// TIA Portal project "SmartFactory_FactoryIO_SortingStation" (V20)

(* hardware
DEVICE "S71500/ET200MP-Station_1"  S7-1500 station
   slot 0: "."  Rack  6ES7 590-1***0-0AA0
   slot 1: "PLC_1"  CPU 1511-1 PN  6ES7 511-1AK02-0AB0  V2.9
      slot 3: "CPU-Display_1"  6ES7591-1AA00-0AA0
      slot 32768: "PLC"  X1
         slot 32769: "Port_1"  X1 P1
         slot 32770: "Port_2"  X1 P2
      slot 34817: "Virtual CP interface port_1"  Virtual CP interface port  Virtual CP interface port
   slot 2: "AI 8xU/I/RTD/TC ST_1"  AI 8xU/I/RTD/TC ST  6ES7 531-7KF00-0AB0  V2.0
   slot 3: "AI 8xU/I/RTD/TC ST_2"  AI 8xU/I/RTD/TC ST  6ES7 531-7KF00-0AB0  V2.0
   slot 4: "AI 8xU/I/RTD/TC ST_3"  AI 8xU/I/RTD/TC ST  6ES7 531-7KF00-0AB0  V2.0
   slot 5: "AI 8xU/I/RTD/TC ST_4"  AI 8xU/I/RTD/TC ST  6ES7 531-7KF00-0AB0  V2.0
   slot 6: "DI 16x24VDC BA_1"  DI 16x24VDC BA  6ES7 521-1BH10-0AA0  V1.0
*)

// ===== PLC "PLC_1"  CPU 1511-1 PN =====

VAR_GLOBAL   // PLC tag table "Standard-Variablentabelle"
   "Start" AT %I0.0 : Bool;
   "Pause & Unpause" AT %I0.1 : Bool;
   "Reset" AT %I0.2 : Bool;
   "Pusher 1 front" AT %I0.3 : Bool;
   "Pusher 2 front" AT %I0.4 : Bool;
   "Pusher 1 back" AT %I0.5 : Bool;
   "Pusher 2 back" AT %I0.6 : Bool;
   "At pusher 1 exit" AT %I0.7 : Bool;
   "At pusher 2 exit" AT %I1.0 : Bool;
   "Sensor 1" AT %I1.1 : Bool;
   "Sensor 2" AT %I1.2 : Bool;
   "Vision sensor 1" AT %ID30 : DInt;
   "Vision sensor 2" AT %ID34 : DInt;
   "Start light" AT %Q0.0 : Bool;
   "P & UP light" AT %Q0.1 : Bool;
   "Reset light" AT %Q0.2 : Bool;
   "Conveyor 1" AT %Q0.3 : Bool;
   "Conveyor 2" AT %Q0.4 : Bool;
   "Entry conveyor 1" AT %Q0.5 : Bool;
   "Entry conveyor 2" AT %Q0.6 : Bool;
   "Pusher 1" AT %Q0.7 : Bool;
   "Pusher 2" AT %Q1.0 : Bool;
   "Blue count" AT %QD30 : DInt;
   "Green count" AT %QD34 : DInt;
   "SYS_RUN_MEM" AT %M0.0 : Bool;
   "SYS_UNPAUSED_MEM" AT %M0.1 : Bool;
   "CASE_C1GREEN_C2BLUE" AT %M0.2 : Bool;
   "GB_ENTRY_CONV1_MEM" AT %M0.3 : Bool;
   "GB_SENSOR1_PULSE_C1" AT %M0.4 : Bool;
   "GB_SENSOR1_NEG_C1" AT %M0.5 : Bool;
   "GB_CONVEYOR1_MEM" AT %M0.6 : Bool;
   "GB_ENTRY_CONV2_MEM" AT %M1.0 : Bool;
   "GB_ATPUSHER2EXIT_NEG_C2" AT %M1.1 : Bool;
   "GB_CONVEYOR2_MEM" AT %M1.2 : Bool;
   "GB_SENSOR1_NEG_P1" AT %M1.3 : Bool;
   "GB_PUSHER1_MEM" AT %M1.4 : Bool;
   "GB_CASE_EXIT" AT %M1.5 : Bool;
   "GB_SENSOR1_NEG_EC1" AT %M1.6 : Bool;
   "GB_ATPUSHER2EXIT_NEG_EC1" AT %M0.7 : Bool;
   "CASE_C1BLUE_C2GREEN" AT %M1.7 : Bool;
   "CASE_BOTH_BLUE" AT %M2.0 : Bool;
   "CASE_BOTH_GREEN" AT %M2.1 : Bool;
   "BG_ENTRY_C1C2_MEM" AT %M2.2 : Bool;
   "BG_CASE_EXIT" AT %M2.3 : Bool;
   "CASE_GB_RESETS_BG_PULSE" AT %M2.4 : Bool;
   "CASE_BG_RESETS_GB_PULSE" AT %M2.5 : Bool;
   "CASE_BB_RESETS_GB_PULSE" AT %M2.6 : Bool;
   "CASE_GG_RESETS_GB_PULSE" AT %M2.7 : Bool;
   "CASE_BB_RESETS_BG_PULSE" AT %M3.0 : Bool;
   "CASE_GG_RESETS_BG_PULSE" AT %M3.1 : Bool;
   "CASE_GB_RESETS_BB_PULSE" AT %M3.2 : Bool;
   "CASE_BG_RESETS_BB_PULSE" AT %M3.3 : Bool;
   "CASE_GG_RESETS_BB_PULSE" AT %M3.4 : Bool;
   "BB_CASE_EXIT" AT %M3.5 : Bool;
   "BB_ENTRY_CONV1_MEM" AT %M3.6 : Bool;
   "BB_CONVEYOR1_MEM" AT %M3.7 : Bool;
   "BB_ENTRY_CONV2_MEM" AT %M4.0 : Bool;
   "BB_CONVEYOR2_MEM" AT %M4.1 : Bool;
   "BB_PUSHER2_MEM" AT %M4.2 : Bool;
   "BB_SENSOR2_NEG" AT %M4.3 : Bool;
   "BB_SENSOR2_PULSE" AT %M4.4 : Bool;
   "BB_SENSOR2_NEG_C2" AT %M4.5 : Bool;
   "BB_SENSOR2_NEG_P2" AT %M4.6 : Bool;
   "BB_ATPUSHER1EXIT_NEG" AT %M4.7 : Bool;
   "BB_ATPUSHER1EXIT_NEG_EC1" AT %M5.0 : Bool;
   "CASE_GB_RESETS_GG_PULSE" AT %M5.1 : Bool;
   "CASE_BG_RESETS_GG_PULSE" AT %M5.2 : Bool;
   "CASE_BB_RESETS_GG_PULSE" AT %M5.3 : Bool;
   "GG_ENTRY_CONV1_MEM" AT %M5.4 : Bool;
   "GG_CONVEYOR1_MEM" AT %M5.5 : Bool;
   "GG_ENTRY_CONV2_MEM" AT %M5.6 : Bool;
   "GG_CONVEYOR2_MEM" AT %M5.7 : Bool;
   "GG_PUSHER1_MEM" AT %M6.0 : Bool;
   "GG_SENSOR1_PULSE" AT %M6.1 : Bool;
   "GG_SENSOR1_NEG_EC1" AT %M6.2 : Bool;
   "GG_SENSOR1_NEG_C1" AT %M6.3 : Bool;
   "GG_SENSOR1_NEG_P1" AT %M6.4 : Bool;
   "GG_ATPUSHER2EXIT_NEG" AT %M6.5 : Bool;
   "GG_ATPUSHER2EXIT_NEG_EC1" AT %M6.6 : Bool;
   "BG_SENSOR1_PULSE" AT %M6.7 : Bool;
   "BG_CONV1CONV2_MEM" AT %M7.0 : Bool;
   "BG_SENSOR1_NEG" AT %M7.1 : Bool;
   "BG_ATPUSHER1EXIT_NEG_C1C2" AT %M7.2 : Bool;
   "BG_ATPUSHER1EXIT_NEG_EC1EC2" AT %M7.3 : Bool;
   "CNT_BLUE_TRIGGER" AT %M7.4 : Bool;
   "CNT_GREEN_TRIGGER" AT %M7.5 : Bool;
   "SYS_PAUSED_MEM" AT %M7.6 : Bool;
END_VAR

// folder: System blocks/Program resources

DATA_BLOCK "IEC_Counter_0_DB"   // DB1
{ S7_Optimized_Access := 'TRUE' }
AUTHOR : SIMATIC
FAMILY : IEC
NAME : DCNTR
VERSION : 1.2
// stored: InstanceOfName IEC_DCOUNTER
"IEC_DCOUNTER"
BEGIN
END_DATA_BLOCK

DATA_BLOCK "IEC_Counter_0_DB_1"   // DB2
{ S7_Optimized_Access := 'TRUE' }
AUTHOR : SIMATIC
FAMILY : IEC
NAME : DCNTR
VERSION : 1.2
// stored: InstanceOfName IEC_DCOUNTER
"IEC_DCOUNTER"
BEGIN
END_DATA_BLOCK

// folder: (top level)

FUNCTION "MHJ-PLC-Lab-Function-S71500" : Void   // FC9000, SCL
{ S7_Optimized_Access := 'TRUE' }
VERSION : 0.1
   VAR_TEMP
      Value : Byte;
      ForCounter : Int;
   END_VAR
   VAR CONSTANT
      Value_01_DW : DWord := 16#1223_5486;
      Value_02_DW : DWord := 16#A6C9_D1F5;
   END_VAR
BEGIN

   #Value:=PEEK(area := 16#82,
        dbNumber := 0,
        byteOffset := 511);
   #Value := #Value + 1;

   POKE(area := 16#82,
        dbNumber := 0,
        byteOffset := 511,
        value := #Value);

   POKE(area := 16#82,
        dbNumber := 0,
        byteOffset := 1016,
        value := #Value_01_DW);
   POKE(area := 16#82,
        dbNumber := 0,
        byteOffset := 1020,
        value := #Value_02_DW);

   FOR #ForCounter := 0 TO 63 DO
       #Value:=PEEK(area := 16#1,
            dbNumber := 0,
            byteOffset := #ForCounter);
       POKE(area := 16#81,
            dbNumber := 0,
            byteOffset := #ForCounter,
            value := #Value);
   END_FOR;
   #Value := PEEK(area := 16#1,
                  dbNumber := 0,
                  byteOffset := 512);
   POKE(area := 16#82,
        dbNumber := 0,
        byteOffset := 512,
        value := #Value);
END_FUNCTION

ORGANIZATION_BLOCK "Main"   // OB1, LAD, ProgramCycle
TITLE = "Main Program Sweep (Cycle)"
{ S7_Optimized_Access := 'TRUE' }
VERSION : 0.1
   VAR_INPUT
      Initial_Call : Bool;   // Initial call of this OB
      Remanence : Bool;   // =True, if remanent data are available
   END_VAR
   VAR_TEMP   // added for the SCL form of the ladder/FBD networks
      _w1 : Bool;
      _w2 : Bool;
      _w3 : Bool;
      _w4 : Bool;
      _w5 : Bool;
      _w6 : Bool;
      _w7 : Bool;
      _w8 : Bool;
      _w9 : Bool;
      _w10 : Bool;
      _w11 : Bool;
      _w12 : Bool;
      _w13 : Bool;
      _w14 : Bool;
   END_VAR
BEGIN

REGION Network 1
   // Lien TIA ↔ Factory I/O (FC9000), ne pas supprimer.
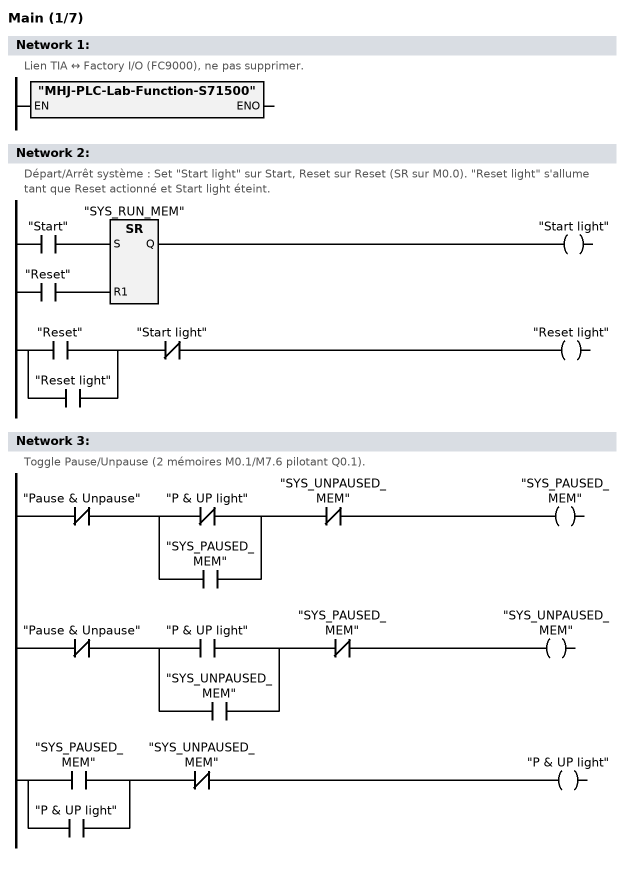
   RUNG wire#powerrail
      "MHJ-PLC-Lab-Function-S71500"()
   END_RUNG
   // the same network as SCL:
   "MHJ-PLC-Lab-Function-S71500"();
END_REGION

REGION Network 2
   // Départ/Arrêt système : Set "Start light" sur Start, Reset sur Reset (SR sur M0.0). "Reset light" s'allume tant que Reset actionné et Start light éteint.
   RUNG wire#powerrail
      Contact( "Start" )
      S_SR(operand := "SYS_RUN_MEM", r1 := wire#w1)
      Coil( "Start light" )
   END_RUNG
   RUNG wire#powerrail
      Contact( "Reset" )
   END_RUNG wire#w1
   RUNG wire#powerrail
      Contact( "Reset" )
      wire#w2
      I_Contact( "Start light" )
      Coil( "Reset light" )
   END_RUNG
   RUNG wire#powerrail
      Contact( "Reset light" )
   END_RUNG wire#w2
   // the same network as SCL:
   IF "Start" THEN
       "SYS_RUN_MEM" := TRUE;   // SR flip-flop
   END_IF;
   IF "Reset" THEN "SYS_RUN_MEM" := FALSE; END_IF;
   "Start light" := "SYS_RUN_MEM";
   "Reset light" := ("Reset" OR "Reset light") AND NOT "Start light";
END_REGION

REGION Network 3
   // Toggle Pause/Unpause (2 mémoires M0.1/M7.6 pilotant Q0.1).
   RUNG wire#powerrail
      I_Contact( "Pause & Unpause" )
      wire#w1
      I_Contact( "P & UP light" )
      wire#w2
      I_Contact( "SYS_UNPAUSED_MEM" )
      Coil( "SYS_PAUSED_MEM" )
   END_RUNG
   RUNG wire#w1
      Contact( "SYS_PAUSED_MEM" )
   END_RUNG wire#w2
   RUNG wire#powerrail
      I_Contact( "Pause & Unpause" )
      wire#w3
      Contact( "P & UP light" )
      wire#w4
      I_Contact( "SYS_PAUSED_MEM" )
      Coil( "SYS_UNPAUSED_MEM" )
   END_RUNG
   RUNG wire#w3
      Contact( "SYS_UNPAUSED_MEM" )
   END_RUNG wire#w4
   RUNG wire#powerrail
      Contact( "SYS_PAUSED_MEM" )
      wire#w5
      I_Contact( "SYS_UNPAUSED_MEM" )
      Coil( "P & UP light" )
   END_RUNG
   RUNG wire#powerrail
      Contact( "P & UP light" )
   END_RUNG wire#w5
   // the same network as SCL:
   "SYS_PAUSED_MEM" := NOT "Pause & Unpause" AND (NOT "P & UP light" OR "SYS_PAUSED_MEM") AND NOT "SYS_UNPAUSED_MEM";
   "SYS_UNPAUSED_MEM" := NOT "Pause & Unpause" AND ("P & UP light" OR "SYS_UNPAUSED_MEM") AND NOT "SYS_PAUSED_MEM";
   "P & UP light" := ("SYS_PAUSED_MEM" OR "P & UP light") AND NOT "SYS_UNPAUSED_MEM";
END_REGION

REGION Network 4
   // Détection de la combinaison couleur des 2 postes (Vision sensor 1=Bleu(1)/Vert(4), idem sensor 2). 4 cas mutuellement exclusifs mémorisés en SR, avec reset croisé par front montant dès qu'un autre cas se déclenche. Comptage Bleu/Vert en sortie (CTU sur "At pusher 1/2 exit").
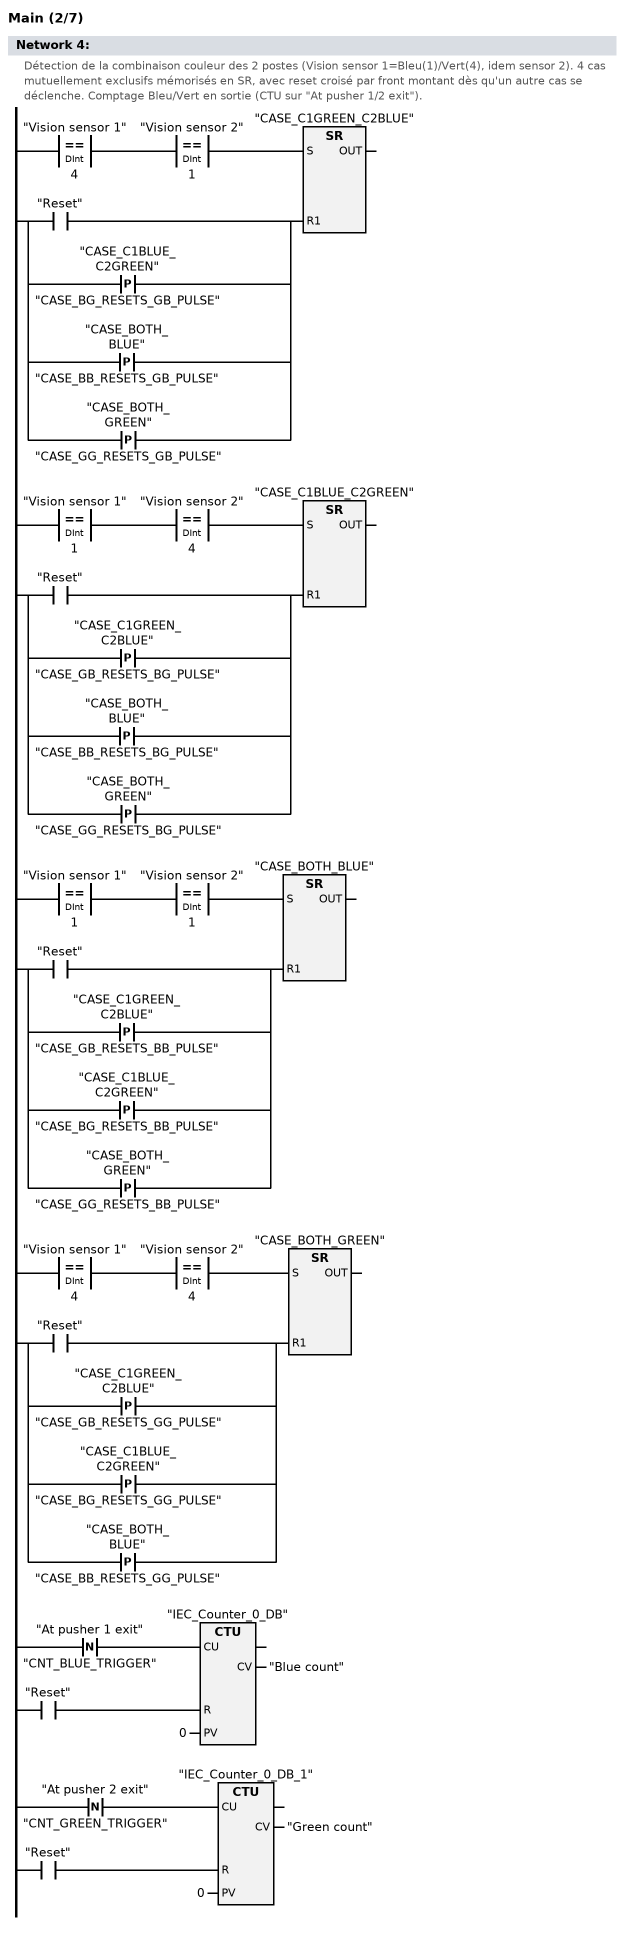
   #_w1 := "CASE_C1BLUE_C2GREEN" AND NOT "CASE_BG_RESETS_GB_PULSE";   // rising edge of "CASE_C1BLUE_C2GREEN"
   "CASE_BG_RESETS_GB_PULSE" := "CASE_C1BLUE_C2GREEN";
   #_w2 := "CASE_BOTH_BLUE" AND NOT "CASE_BB_RESETS_GB_PULSE";   // rising edge of "CASE_BOTH_BLUE"
   "CASE_BB_RESETS_GB_PULSE" := "CASE_BOTH_BLUE";
   #_w3 := "CASE_BOTH_GREEN" AND NOT "CASE_GG_RESETS_GB_PULSE";   // rising edge of "CASE_BOTH_GREEN"
   "CASE_GG_RESETS_GB_PULSE" := "CASE_BOTH_GREEN";
   IF ("Vision sensor 1" = 4) AND ("Vision sensor 2" = 1) THEN
       "CASE_C1GREEN_C2BLUE" := TRUE;   // SR flip-flop
   END_IF;
   IF "Reset" OR #_w1 OR #_w2 OR #_w3 THEN "CASE_C1GREEN_C2BLUE" := FALSE; END_IF;
   #_w4 := "CASE_C1GREEN_C2BLUE" AND NOT "CASE_GB_RESETS_BG_PULSE";   // rising edge of "CASE_C1GREEN_C2BLUE"
   "CASE_GB_RESETS_BG_PULSE" := "CASE_C1GREEN_C2BLUE";
   #_w5 := "CASE_BOTH_BLUE" AND NOT "CASE_BB_RESETS_BG_PULSE";   // rising edge of "CASE_BOTH_BLUE"
   "CASE_BB_RESETS_BG_PULSE" := "CASE_BOTH_BLUE";
   #_w6 := "CASE_BOTH_GREEN" AND NOT "CASE_GG_RESETS_BG_PULSE";   // rising edge of "CASE_BOTH_GREEN"
   "CASE_GG_RESETS_BG_PULSE" := "CASE_BOTH_GREEN";
   IF ("Vision sensor 1" = 1) AND ("Vision sensor 2" = 4) THEN
       "CASE_C1BLUE_C2GREEN" := TRUE;   // SR flip-flop
   END_IF;
   IF "Reset" OR #_w4 OR #_w5 OR #_w6 THEN "CASE_C1BLUE_C2GREEN" := FALSE; END_IF;
   #_w7 := "CASE_C1GREEN_C2BLUE" AND NOT "CASE_GB_RESETS_BB_PULSE";   // rising edge of "CASE_C1GREEN_C2BLUE"
   "CASE_GB_RESETS_BB_PULSE" := "CASE_C1GREEN_C2BLUE";
   #_w8 := "CASE_C1BLUE_C2GREEN" AND NOT "CASE_BG_RESETS_BB_PULSE";   // rising edge of "CASE_C1BLUE_C2GREEN"
   "CASE_BG_RESETS_BB_PULSE" := "CASE_C1BLUE_C2GREEN";
   #_w9 := "CASE_BOTH_GREEN" AND NOT "CASE_GG_RESETS_BB_PULSE";   // rising edge of "CASE_BOTH_GREEN"
   "CASE_GG_RESETS_BB_PULSE" := "CASE_BOTH_GREEN";
   IF ("Vision sensor 1" = 1) AND ("Vision sensor 2" = 1) THEN
       "CASE_BOTH_BLUE" := TRUE;   // SR flip-flop
   END_IF;
   IF "Reset" OR #_w7 OR #_w8 OR #_w9 THEN "CASE_BOTH_BLUE" := FALSE; END_IF;
   #_w10 := "CASE_C1GREEN_C2BLUE" AND NOT "CASE_GB_RESETS_GG_PULSE";   // rising edge of "CASE_C1GREEN_C2BLUE"
   "CASE_GB_RESETS_GG_PULSE" := "CASE_C1GREEN_C2BLUE";
   #_w11 := "CASE_C1BLUE_C2GREEN" AND NOT "CASE_BG_RESETS_GG_PULSE";   // rising edge of "CASE_C1BLUE_C2GREEN"
   "CASE_BG_RESETS_GG_PULSE" := "CASE_C1BLUE_C2GREEN";
   #_w12 := "CASE_BOTH_BLUE" AND NOT "CASE_BB_RESETS_GG_PULSE";   // rising edge of "CASE_BOTH_BLUE"
   "CASE_BB_RESETS_GG_PULSE" := "CASE_BOTH_BLUE";
   IF ("Vision sensor 1" = 4) AND ("Vision sensor 2" = 4) THEN
       "CASE_BOTH_GREEN" := TRUE;   // SR flip-flop
   END_IF;
   IF "Reset" OR #_w10 OR #_w11 OR #_w12 THEN "CASE_BOTH_GREEN" := FALSE; END_IF;
   #_w13 := NOT "At pusher 1 exit" AND "CNT_BLUE_TRIGGER";   // falling edge of "At pusher 1 exit"
   "CNT_BLUE_TRIGGER" := "At pusher 1 exit";
   "IEC_Counter_0_DB".CTU(CU := #_w13, R := "Reset", PV := 0, CV => "Blue count");
   #_w14 := NOT "At pusher 2 exit" AND "CNT_GREEN_TRIGGER";   // falling edge of "At pusher 2 exit"
   "CNT_GREEN_TRIGGER" := "At pusher 2 exit";
   "IEC_Counter_0_DB_1".CTU(CU := #_w14, R := "Reset", PV := 0, CV => "Green count");
END_REGION

REGION Network 5
   // Si le cas "Vert sur Conv1 / Bleu sur Conv2" est actif → saut vers Network 9, les Networks 10 à 12 sont ignorés ce cycle.
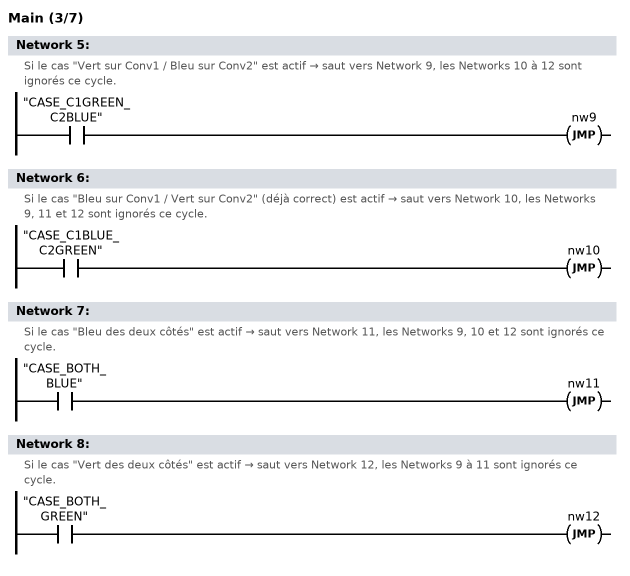
   RUNG wire#powerrail
      Contact( "CASE_C1GREEN_C2BLUE" )
      JumpCoil( nw9 )
   END_RUNG
   // the same network as SCL:
   IF "CASE_C1GREEN_C2BLUE" THEN GOTO nw9; END_IF;
END_REGION

REGION Network 6
   // Si le cas "Bleu sur Conv1 / Vert sur Conv2" (déjà correct) est actif → saut vers Network 10, les Networks 9, 11 et 12 sont ignorés ce cycle.
   RUNG wire#powerrail
      Contact( "CASE_C1BLUE_C2GREEN" )
      JumpCoil( nw10 )
   END_RUNG
   // the same network as SCL:
   IF "CASE_C1BLUE_C2GREEN" THEN GOTO nw10; END_IF;
END_REGION

REGION Network 7
   // Si le cas "Bleu des deux côtés" est actif → saut vers Network 11, les Networks 9, 10 et 12 sont ignorés ce cycle.
   RUNG wire#powerrail
      Contact( "CASE_BOTH_BLUE" )
      JumpCoil( nw11 )
   END_RUNG
   // the same network as SCL:
   IF "CASE_BOTH_BLUE" THEN GOTO nw11; END_IF;
END_REGION

REGION Network 8
   // Si le cas "Vert des deux côtés" est actif → saut vers Network 12, les Networks 9 à 11 sont ignorés ce cycle.
   RUNG wire#powerrail
      Contact( "CASE_BOTH_GREEN" )
      JumpCoil( nw12 )
   END_RUNG
   // the same network as SCL:
   IF "CASE_BOTH_GREEN" THEN GOTO nw12; END_IF;
END_REGION

REGION Network 9
   // Cas Vert/Bleu (positions inversées) : active les 2 convoyeurs d'entrée + convoyeur 1 sur détection Sensor 1, puis Pousseur 1 transfère l'objet Vert du convoyeur 1 vers le convoyeur 2 dès qu'il atteint la butée. RET dès que le cas GB n'est plus actif.
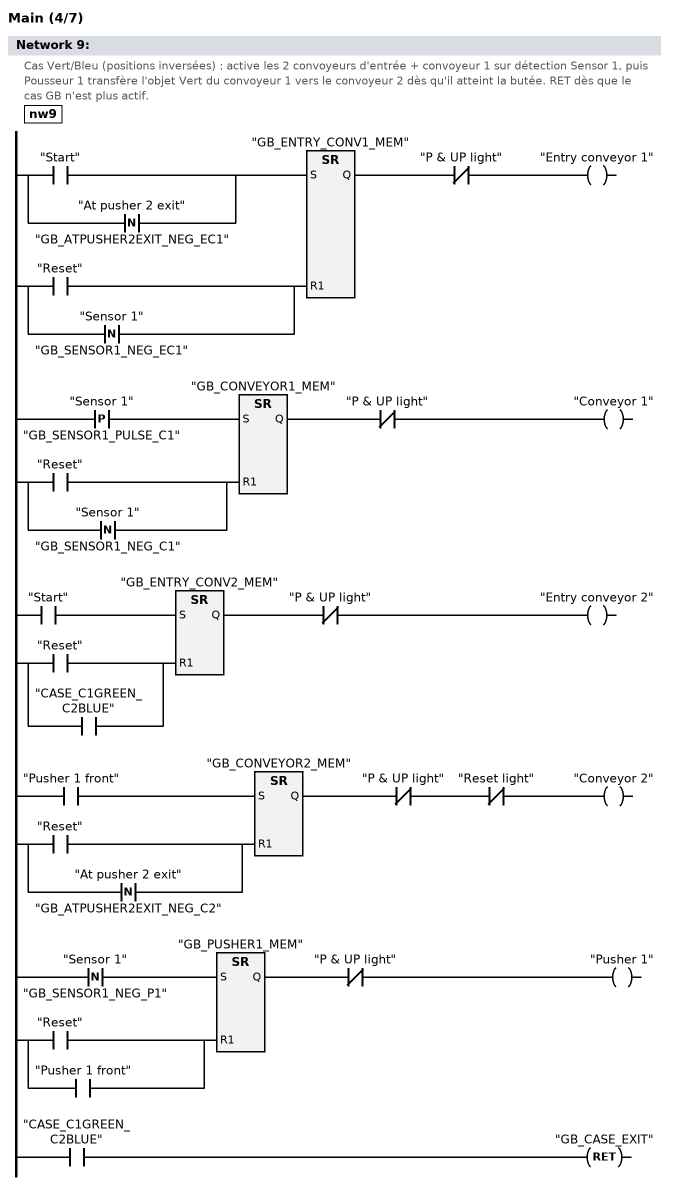
   nw9:
   #_w1 := NOT "At pusher 2 exit" AND "GB_ATPUSHER2EXIT_NEG_EC1";   // falling edge of "At pusher 2 exit"
   "GB_ATPUSHER2EXIT_NEG_EC1" := "At pusher 2 exit";
   #_w2 := NOT "Sensor 1" AND "GB_SENSOR1_NEG_EC1";   // falling edge of "Sensor 1"
   "GB_SENSOR1_NEG_EC1" := "Sensor 1";
   IF "Start" OR #_w1 THEN
       "GB_ENTRY_CONV1_MEM" := TRUE;   // SR flip-flop
   END_IF;
   IF "Reset" OR #_w2 THEN "GB_ENTRY_CONV1_MEM" := FALSE; END_IF;
   "Entry conveyor 1" := "GB_ENTRY_CONV1_MEM" AND NOT "P & UP light";
   #_w3 := "Sensor 1" AND NOT "GB_SENSOR1_PULSE_C1";   // rising edge of "Sensor 1"
   "GB_SENSOR1_PULSE_C1" := "Sensor 1";
   #_w4 := NOT "Sensor 1" AND "GB_SENSOR1_NEG_C1";   // falling edge of "Sensor 1"
   "GB_SENSOR1_NEG_C1" := "Sensor 1";
   IF #_w3 THEN
       "GB_CONVEYOR1_MEM" := TRUE;   // SR flip-flop
   END_IF;
   IF "Reset" OR #_w4 THEN "GB_CONVEYOR1_MEM" := FALSE; END_IF;
   "Conveyor 1" := "GB_CONVEYOR1_MEM" AND NOT "P & UP light";
   IF "Start" THEN
       "GB_ENTRY_CONV2_MEM" := TRUE;   // SR flip-flop
   END_IF;
   IF "Reset" OR "CASE_C1GREEN_C2BLUE" THEN "GB_ENTRY_CONV2_MEM" := FALSE; END_IF;
   "Entry conveyor 2" := "GB_ENTRY_CONV2_MEM" AND NOT "P & UP light";
   #_w5 := NOT "At pusher 2 exit" AND "GB_ATPUSHER2EXIT_NEG_C2";   // falling edge of "At pusher 2 exit"
   "GB_ATPUSHER2EXIT_NEG_C2" := "At pusher 2 exit";
   IF "Pusher 1 front" THEN
       "GB_CONVEYOR2_MEM" := TRUE;   // SR flip-flop
   END_IF;
   IF "Reset" OR #_w5 THEN "GB_CONVEYOR2_MEM" := FALSE; END_IF;
   "Conveyor 2" := "GB_CONVEYOR2_MEM" AND NOT "P & UP light" AND NOT "Reset light";
   #_w6 := NOT "Sensor 1" AND "GB_SENSOR1_NEG_P1";   // falling edge of "Sensor 1"
   "GB_SENSOR1_NEG_P1" := "Sensor 1";
   IF #_w6 THEN
       "GB_PUSHER1_MEM" := TRUE;   // SR flip-flop
   END_IF;
   IF "Reset" OR "Pusher 1 front" THEN "GB_PUSHER1_MEM" := FALSE; END_IF;
   "Pusher 1" := "GB_PUSHER1_MEM" AND NOT "P & UP light";
   IF "CASE_C1GREEN_C2BLUE" THEN
       ENO := "GB_CASE_EXIT";
       RETURN;
   END_IF;
END_REGION

REGION Network 10
   // Cas Bleu/Vert déjà en bonne position : active simplement les 2 convoyeurs d'entrée + les 2 convoyeurs principaux, aucun pousseur nécessaire.
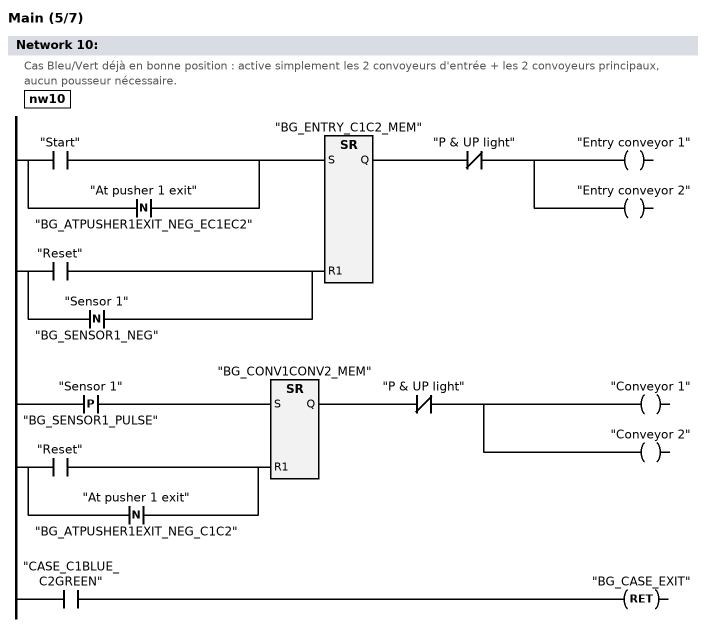
   nw10:
   #_w1 := NOT "At pusher 1 exit" AND "BG_ATPUSHER1EXIT_NEG_EC1EC2";   // falling edge of "At pusher 1 exit"
   "BG_ATPUSHER1EXIT_NEG_EC1EC2" := "At pusher 1 exit";
   #_w2 := NOT "Sensor 1" AND "BG_SENSOR1_NEG";   // falling edge of "Sensor 1"
   "BG_SENSOR1_NEG" := "Sensor 1";
   IF "Start" OR #_w1 THEN
       "BG_ENTRY_C1C2_MEM" := TRUE;   // SR flip-flop
   END_IF;
   IF "Reset" OR #_w2 THEN "BG_ENTRY_C1C2_MEM" := FALSE; END_IF;
   "Entry conveyor 1" := "BG_ENTRY_C1C2_MEM" AND NOT "P & UP light";
   "Entry conveyor 2" := "Entry conveyor 1";
   #_w3 := "Sensor 1" AND NOT "BG_SENSOR1_PULSE";   // rising edge of "Sensor 1"
   "BG_SENSOR1_PULSE" := "Sensor 1";
   #_w4 := NOT "At pusher 1 exit" AND "BG_ATPUSHER1EXIT_NEG_C1C2";   // falling edge of "At pusher 1 exit"
   "BG_ATPUSHER1EXIT_NEG_C1C2" := "At pusher 1 exit";
   IF #_w3 THEN
       "BG_CONV1CONV2_MEM" := TRUE;   // SR flip-flop
   END_IF;
   IF "Reset" OR #_w4 THEN "BG_CONV1CONV2_MEM" := FALSE; END_IF;
   "Conveyor 1" := "BG_CONV1CONV2_MEM" AND NOT "P & UP light";
   "Conveyor 2" := "Conveyor 1";
   IF "CASE_C1BLUE_C2GREEN" THEN
       ENO := "BG_CASE_EXIT";
       RETURN;
   END_IF;
END_REGION

REGION Network 11
   // Cas Bleu des deux côtés : Pousseur 2 renvoie l'objet Bleu en excès du convoyeur 2 vers le convoyeur 1 (symétrique de N9, sur Sensor 2/Pousseur 2).
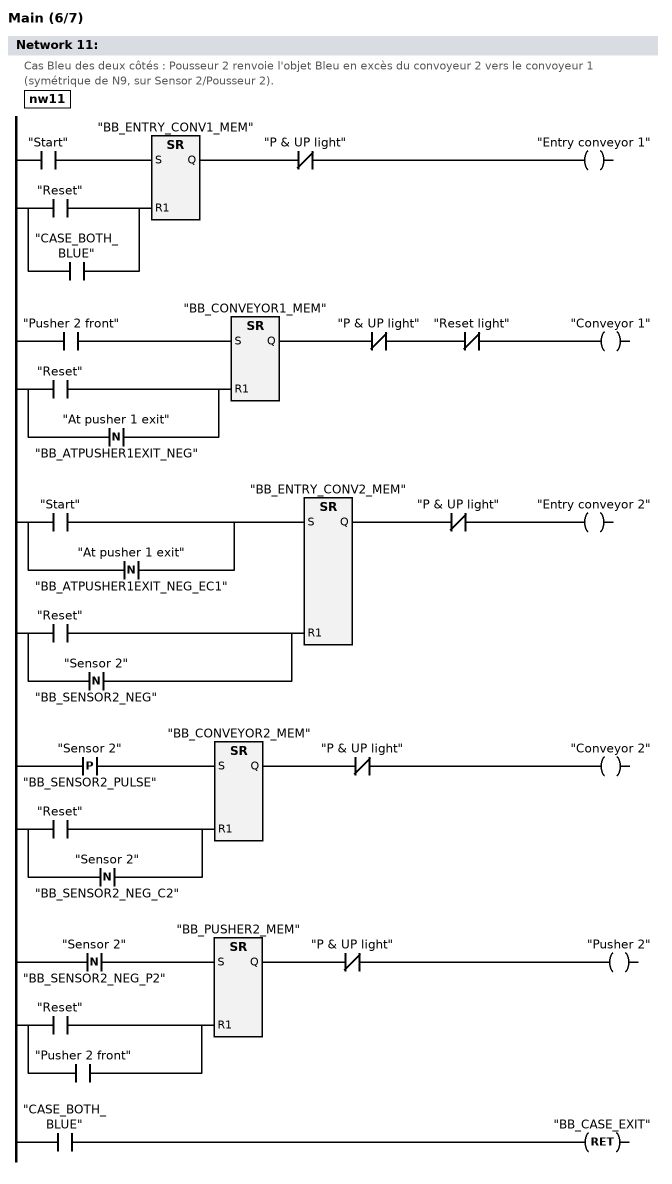
   nw11:
   IF "Start" THEN
       "BB_ENTRY_CONV1_MEM" := TRUE;   // SR flip-flop
   END_IF;
   IF "Reset" OR "CASE_BOTH_BLUE" THEN "BB_ENTRY_CONV1_MEM" := FALSE; END_IF;
   "Entry conveyor 1" := "BB_ENTRY_CONV1_MEM" AND NOT "P & UP light";
   #_w1 := NOT "At pusher 1 exit" AND "BB_ATPUSHER1EXIT_NEG";   // falling edge of "At pusher 1 exit"
   "BB_ATPUSHER1EXIT_NEG" := "At pusher 1 exit";
   IF "Pusher 2 front" THEN
       "BB_CONVEYOR1_MEM" := TRUE;   // SR flip-flop
   END_IF;
   IF "Reset" OR #_w1 THEN "BB_CONVEYOR1_MEM" := FALSE; END_IF;
   "Conveyor 1" := "BB_CONVEYOR1_MEM" AND NOT "P & UP light" AND NOT "Reset light";
   #_w2 := NOT "At pusher 1 exit" AND "BB_ATPUSHER1EXIT_NEG_EC1";   // falling edge of "At pusher 1 exit"
   "BB_ATPUSHER1EXIT_NEG_EC1" := "At pusher 1 exit";
   #_w3 := NOT "Sensor 2" AND "BB_SENSOR2_NEG";   // falling edge of "Sensor 2"
   "BB_SENSOR2_NEG" := "Sensor 2";
   IF "Start" OR #_w2 THEN
       "BB_ENTRY_CONV2_MEM" := TRUE;   // SR flip-flop
   END_IF;
   IF "Reset" OR #_w3 THEN "BB_ENTRY_CONV2_MEM" := FALSE; END_IF;
   "Entry conveyor 2" := "BB_ENTRY_CONV2_MEM" AND NOT "P & UP light";
   #_w4 := "Sensor 2" AND NOT "BB_SENSOR2_PULSE";   // rising edge of "Sensor 2"
   "BB_SENSOR2_PULSE" := "Sensor 2";
   #_w5 := NOT "Sensor 2" AND "BB_SENSOR2_NEG_C2";   // falling edge of "Sensor 2"
   "BB_SENSOR2_NEG_C2" := "Sensor 2";
   IF #_w4 THEN
       "BB_CONVEYOR2_MEM" := TRUE;   // SR flip-flop
   END_IF;
   IF "Reset" OR #_w5 THEN "BB_CONVEYOR2_MEM" := FALSE; END_IF;
   "Conveyor 2" := "BB_CONVEYOR2_MEM" AND NOT "P & UP light";
   #_w6 := NOT "Sensor 2" AND "BB_SENSOR2_NEG_P2";   // falling edge of "Sensor 2"
   "BB_SENSOR2_NEG_P2" := "Sensor 2";
   IF #_w6 THEN
       "BB_PUSHER2_MEM" := TRUE;   // SR flip-flop
   END_IF;
   IF "Reset" OR "Pusher 2 front" THEN "BB_PUSHER2_MEM" := FALSE; END_IF;
   "Pusher 2" := "BB_PUSHER2_MEM" AND NOT "P & UP light";
   IF "CASE_BOTH_BLUE" THEN
       ENO := "BB_CASE_EXIT";
       RETURN;
   END_IF;
END_REGION

REGION Network 12
   // Cas Vert des deux côtés : Pousseur 1 déplace l'objet Vert en excès du convoyeur 1 vers le convoyeur 2 (même logique que N9).
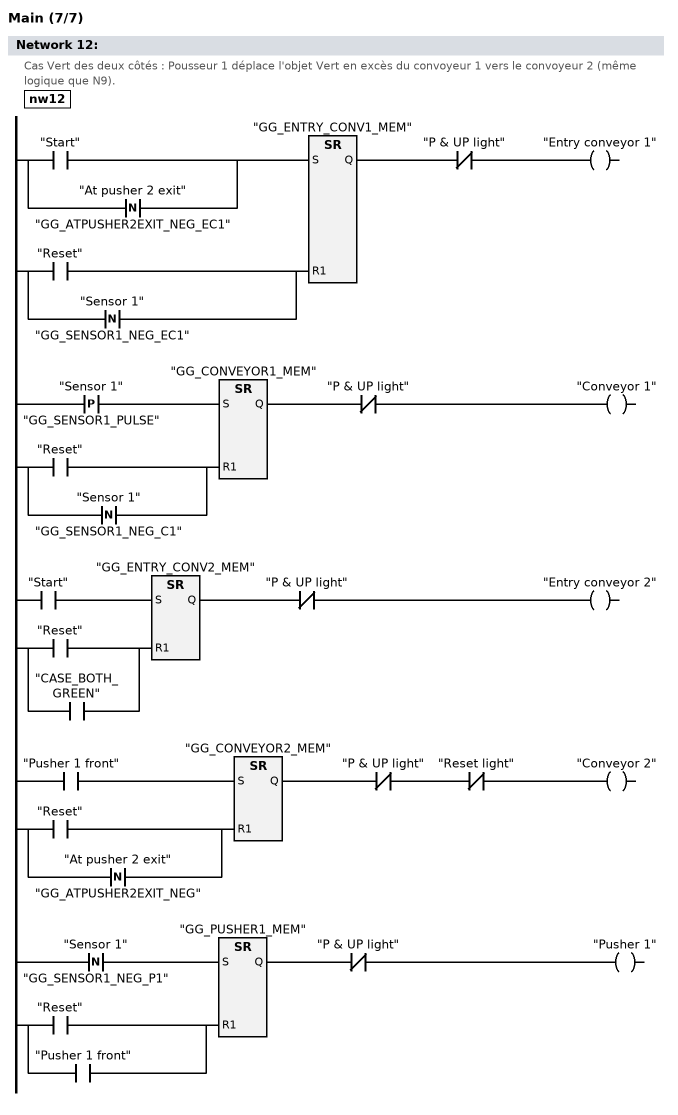
   Label( nw12 )
   RUNG wire#powerrail
      Contact( "Start" )
      wire#w1
      S_SR(operand := "GG_ENTRY_CONV1_MEM", r1 := wire#w2)
      I_Contact( "P & UP light" )
      Coil( "Entry conveyor 1" )
   END_RUNG
   RUNG wire#powerrail
      N_Contact(operand := "At pusher 2 exit", bit := "GG_ATPUSHER2EXIT_NEG_EC1")
   END_RUNG wire#w1
   RUNG wire#powerrail
      Contact( "Reset" )
   END_RUNG wire#w2
   RUNG wire#powerrail
      N_Contact(operand := "Sensor 1", bit := "GG_SENSOR1_NEG_EC1")
   END_RUNG wire#w2
   RUNG wire#powerrail
      P_Contact(operand := "Sensor 1", bit := "GG_SENSOR1_PULSE")
      S_SR(operand := "GG_CONVEYOR1_MEM", r1 := wire#w3)
      I_Contact( "P & UP light" )
      Coil( "Conveyor 1" )
   END_RUNG
   RUNG wire#powerrail
      Contact( "Reset" )
   END_RUNG wire#w3
   RUNG wire#powerrail
      N_Contact(operand := "Sensor 1", bit := "GG_SENSOR1_NEG_C1")
   END_RUNG wire#w3
   RUNG wire#powerrail
      Contact( "Start" )
      S_SR(operand := "GG_ENTRY_CONV2_MEM", r1 := wire#w4)
      I_Contact( "P & UP light" )
      Coil( "Entry conveyor 2" )
   END_RUNG
   RUNG wire#powerrail
      Contact( "Reset" )
   END_RUNG wire#w4
   RUNG wire#powerrail
      Contact( "CASE_BOTH_GREEN" )
   END_RUNG wire#w4
   RUNG wire#powerrail
      Contact( "Pusher 1 front" )
      S_SR(operand := "GG_CONVEYOR2_MEM", r1 := wire#w5)
      I_Contact( "P & UP light" )
      I_Contact( "Reset light" )
      Coil( "Conveyor 2" )
   END_RUNG
   RUNG wire#powerrail
      Contact( "Reset" )
   END_RUNG wire#w5
   RUNG wire#powerrail
      N_Contact(operand := "At pusher 2 exit", bit := "GG_ATPUSHER2EXIT_NEG")
   END_RUNG wire#w5
   RUNG wire#powerrail
      N_Contact(operand := "Sensor 1", bit := "GG_SENSOR1_NEG_P1")
      S_SR(operand := "GG_PUSHER1_MEM", r1 := wire#w6)
      I_Contact( "P & UP light" )
      Coil( "Pusher 1" )
   END_RUNG
   RUNG wire#powerrail
      Contact( "Reset" )
   END_RUNG wire#w6
   RUNG wire#powerrail
      Contact( "Pusher 1 front" )
   END_RUNG wire#w6
   // the same network as SCL:
   nw12:
   #_w1 := NOT "At pusher 2 exit" AND "GG_ATPUSHER2EXIT_NEG_EC1";   // falling edge of "At pusher 2 exit"
   "GG_ATPUSHER2EXIT_NEG_EC1" := "At pusher 2 exit";
   #_w2 := NOT "Sensor 1" AND "GG_SENSOR1_NEG_EC1";   // falling edge of "Sensor 1"
   "GG_SENSOR1_NEG_EC1" := "Sensor 1";
   IF "Start" OR #_w1 THEN
       "GG_ENTRY_CONV1_MEM" := TRUE;   // SR flip-flop
   END_IF;
   IF "Reset" OR #_w2 THEN "GG_ENTRY_CONV1_MEM" := FALSE; END_IF;
   "Entry conveyor 1" := "GG_ENTRY_CONV1_MEM" AND NOT "P & UP light";
   #_w3 := "Sensor 1" AND NOT "GG_SENSOR1_PULSE";   // rising edge of "Sensor 1"
   "GG_SENSOR1_PULSE" := "Sensor 1";
   #_w4 := NOT "Sensor 1" AND "GG_SENSOR1_NEG_C1";   // falling edge of "Sensor 1"
   "GG_SENSOR1_NEG_C1" := "Sensor 1";
   IF #_w3 THEN
       "GG_CONVEYOR1_MEM" := TRUE;   // SR flip-flop
   END_IF;
   IF "Reset" OR #_w4 THEN "GG_CONVEYOR1_MEM" := FALSE; END_IF;
   "Conveyor 1" := "GG_CONVEYOR1_MEM" AND NOT "P & UP light";
   IF "Start" THEN
       "GG_ENTRY_CONV2_MEM" := TRUE;   // SR flip-flop
   END_IF;
   IF "Reset" OR "CASE_BOTH_GREEN" THEN "GG_ENTRY_CONV2_MEM" := FALSE; END_IF;
   "Entry conveyor 2" := "GG_ENTRY_CONV2_MEM" AND NOT "P & UP light";
   #_w5 := NOT "At pusher 2 exit" AND "GG_ATPUSHER2EXIT_NEG";   // falling edge of "At pusher 2 exit"
   "GG_ATPUSHER2EXIT_NEG" := "At pusher 2 exit";
   IF "Pusher 1 front" THEN
       "GG_CONVEYOR2_MEM" := TRUE;   // SR flip-flop
   END_IF;
   IF "Reset" OR #_w5 THEN "GG_CONVEYOR2_MEM" := FALSE; END_IF;
   "Conveyor 2" := "GG_CONVEYOR2_MEM" AND NOT "P & UP light" AND NOT "Reset light";
   #_w6 := NOT "Sensor 1" AND "GG_SENSOR1_NEG_P1";   // falling edge of "Sensor 1"
   "GG_SENSOR1_NEG_P1" := "Sensor 1";
   IF #_w6 THEN
       "GG_PUSHER1_MEM" := TRUE;   // SR flip-flop
   END_IF;
   IF "Reset" OR "Pusher 1 front" THEN "GG_PUSHER1_MEM" := FALSE; END_IF;
   "Pusher 1" := "GG_PUSHER1_MEM" AND NOT "P & UP light";
END_REGION
END_ORGANIZATION_BLOCK